(* CODESYS project settings.library
   DefaultNamespace: KOSTAL.AF2024.Core.Settings
   DocFormat: reStructuredText
   Description: base settings
   Author: Frank Dümpelmann
   Title: KOSTAL.AF2024.Core.Settings
   Version: 1.0.0.0
   Company: KOSTAL GmbH & Co.KG
   Placeholder: KOSTAL.AF2024.Core.Settings

Project tree, tasks and I/O mapping:
  Project Information/
    function F_GetCompany [ST]
    function F_GetTitle [ST]
    function F_GetVersion [ST]
  Version/
    global variables Global_Version
  global variables GVL_CONSTANT
  data type T_MaxString
  data type T_MaxString_UTF8
*)

// T_MaxString
TYPE T_MaxString : WSTRING(255); END_TYPE

// T_MaxString_UTF8
TYPE T_MaxString_UTF8 : STRING(255); END_TYPE

// Version/Global_Version
{attribute 'TcGenerated'}
{attribute 'no-analysis'}
{attribute 'linkalways'}
// This function has been automatically generated from the project information.
VAR_GLOBAL CONSTANT
	{attribute 'const_non_replaced'}
	stLibVersion_KOSTAL_AF2024_Core_Settings : ST_LibVersion := (iMajor := 1, iMinor := 0, iBuild := 0, iRevision := 0, nFlags := 0, sVersion := '1.0.0.0');
END_VAR

// GVL_CONSTANT
{attribute 'qualified_only'}
VAR_GLOBAL CONSTANT
	UNICODE_BigEndian			: WORD:= 16#FFFF;
	UNICODE_LittleEndian	: WORD:= 16#FEFE;
END_VAR

// Project Information/F_GetCompany
// This function has been automatically generated from the project information.
{attribute 'signature_flag' := '1073741824'}
{attribute 'TcGenerated'}
{attribute 'no-analysis'}
FUNCTION F_GetCompany : WSTRING
VAR_INPUT
	
END_VAR

F_GetCompany := "KOSTAL GmbH & Co.KG";

END_FUNCTION

// Project Information/F_GetTitle
// This function has been automatically generated from the project information.
{attribute 'signature_flag' := '1073741824'}
{attribute 'TcGenerated'}
{attribute 'no-analysis'}
FUNCTION F_GetTitle : WSTRING
VAR_INPUT
	
END_VAR

F_GetTitle := "KOSTAL.AF2024.Core.Settings";

END_FUNCTION

// Project Information/F_GetVersion
// This function has been automatically generated from the project information.
{attribute 'signature_flag' := '1073741824'}
{attribute 'TcGenerated'}
{attribute 'no-analysis'}
FUNCTION F_GetVersion : ST_LibVersion
VAR_INPUT
	
END_VAR

F_GetVersion.iMajor := 1;
F_GetVersion.iMinor := 0;
F_GetVersion.iBuild := 0;
F_GetVersion.iRevision := 0;
F_GetVersion.sVersion := '1.0.0.0';
F_GetVersion.nFlags := 0;

END_FUNCTION
